Staubli VAL3: HMI_safezone.dtx

mdesc mNomSpeed = {blend=off}
string sList
string sSelZone
bool bSetFrame
bool bTeach1
bool bMove
bool bRename
bool bConfirm
bool bActive
public num nFrame[6]
num nTRSF1[6]
num nTRSF2[6]
string sLastZone
num _nZoneIndex
string sComment
frame fFrame = {fatherId=world[0]}
bool bBack
tool tTool = {fatherId=flange[0]}
bool bSetFrameData
string sToolIndex
